{attribute 'qualified_only'}
{attribute 'strict'}
{attribute 'to_string'}
TYPE E_Byte :
(
	eOptionA := 0,
	eOptionB,
	eOptionC
) BYTE;
END_TYPE

(* stored: Version 1.1.0.1, ProductVersion 3.1.4026.19
   DUT E_Byte: Id {ffb05ed2-ab96-4dcc-9eed-85de04d21c46} *)
